(* IEC 61131-3 sources: rusty/compiler/plc_cfc/fixtures/blocks/valid/program_negated, 1 file *)

(* ---- program_0.st ---- *)
PROGRAM program_0
VAR_INPUT
    in : DINT;
END_VAR
VAR_IN_OUT
    inout : DINT;
END_VAR
VAR_OUTPUT
    out : DINT;
END_VAR
    out := in + inout;
END_PROGRAM
